PROGRAM Gr01Simulation
VAR_INPUT
	(* Input variables / Eingang Variablen *)
	bEnable								:BOOL;						(* Enable Gr05Persistent *)
END_VAR
VAR
	(* Enummerations *)

	(* Variables *)

	(* References *)

	(* Interfaces *)

	(* Instances *)
END_VAR

IF NOT bEnable
THEN

	RETURN;
END_IF;

A_ForceInput();

ACTION A_ForceInput:


GVL_Gr00IO.binGr00AirPressureOK := TRUE;
GVL_Gr00IO.binGr00LightCurtainOK := TRUE;
GVL_Gr00IO.arbinGr00PowerSupplyOn[2] := TRUE;
GVL_Gr00IO.arbinGr00PowerSupplyOn[3] := TRUE;
GVL_Gr00IO.arbinGr00PowerSupplyOn[4] := TRUE;
GVL_Gr00IO.arbinGr00PowerSupplyOn[5] := TRUE;
GVL_Gr00IO.arbinGr00DoorsClosed[1] := TRUE;
GVL_Gr00IO.arbinGr00DoorsClosed[2] := TRUE;
GVL_Gr00IO.arbinGr00DoorsClosed[3] := TRUE;
GVL_Gr00IO.arbinGr00DoorsClosed[4] := TRUE;
GVL_Gr00IO.arbinGr00DoorsClosed[5] := TRUE;
GVL_Gr00IO.binGr00AllDoorsClosed := GVL_Gr00IO.arbinGr00DoorsClosed[1]
								AND GVL_Gr00IO.arbinGr00DoorsClosed[2]
								AND GVL_Gr00IO.arbinGr00DoorsClosed[3]
								AND GVL_Gr00IO.arbinGr00DoorsClosed[4]
								AND GVL_Gr00IO.arbinGr00DoorsClosed[5];

GVL_Gr00IO.binGr00AllDoorsLocked := TRUE;
GVL_Gr00IO.binGr00TempOK := TRUE;


// only for simulation
// GVL_Gr00IO.binNoEmergencyStop := TRUE;
// GVL_Gr00IO.binMoveRelease := TRUE;
// GVL_Gr00IO.binMoveReleaseSB := TRUE;
END_ACTION

END_PROGRAM

(* stored: Version 1.1.0.1, ProductVersion 3.1.4024.15
   POU Gr01Simulation: Id {86f70c82-c969-4145-a51e-2780e87c2377}, SpecialFunc None
   Action A_ForceInput: Id {3791caab-563f-44be-9114-ddb22f78ffc2} *)
